Fanuc KAREL source: ko00108.KL

-- PROVISIONAL review KL for V770-1; original PC SHA256 b05d4ced9f50d276c5c8dd84dbcf790411ec813109ccf0bb9dd9321a58c336eb
-- Incomplete behavior may be omitted. Consult companion uncertainty JSON. Do not deploy.
PROGRAM KO00108
%NOLOCKGROUP
VAR
  A : REAL
  B : REAL
  OUT : REAL
BEGIN
  -- UNRESOLVED_PC offsets 5-13; opcodes 9D,64,23
  -- UNRESOLVED_PC offsets 18-30; opcodes 2E,64,23
  -- UNRESOLVED_PC offsets 35-56; opcodes 27,22,22,76,23
  -- UNRESOLVED_PC offsets 61-65; opcodes 7F
END KO00108
